SUBAPPLICATION Sitzventile (* Subapplication Type *)
  (* Standard: 61499-2 *)
  (* Version 1.0, 2023-02-11, franz *)
  IMPORT DataPanel::io::MI::DQ::DataPanel_MI_DO::Invalid;
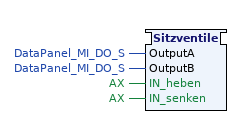
  VAR_INPUT
    OutputA : DataPanel::io::MI::DQ::DataPanel_MI_DO_S := Invalid;
    OutputB : DataPanel::io::MI::DQ::DataPanel_MI_DO_S := Invalid;
  END_VAR
  SOCKETS
    IN_heben : adapter::types::unidirectional::AX;
    IN_senken : adapter::types::unidirectional::AX;
  END_SOCKETS
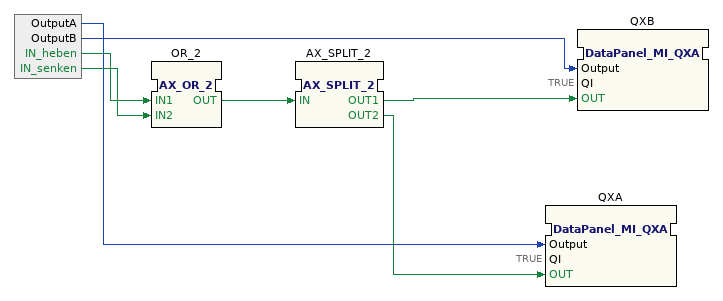
  FBS
    OR_2 : adapter::booleanOperators::AX_OR_2;
    AX_SPLIT_2 : adapter::events::unidirectional::AX_SPLIT_2;
    QXB : DataPanel::io::MI::DQ::DataPanel_MI_QXA(QI := TRUE);
    QXA : DataPanel::io::MI::DQ::DataPanel_MI_QXA(QI := TRUE);
  END_FBS
  DATA_CONNECTIONS
    OutputB TO QXB.Output;
    OutputA TO QXA.Output;
  END_CONNECTIONS
  ADAPTER_CONNECTIONS
    IN_heben TO OR_2.IN1;
    IN_senken TO OR_2.IN2;
    OR_2.OUT TO AX_SPLIT_2.IN;
    AX_SPLIT_2.OUT1 TO QXB.OUT;
    AX_SPLIT_2.OUT2 TO QXA.OUT;
  END_CONNECTIONS
END_SUBAPPLICATION
